(* IEC 61131-3 sources: Versio-VersionControlSystem/fixtures/projects/TC3_PlcSample_reStrText/TC3_PlcSample_reStrText/LibraryDocumentationSample Project/LibPOUs/B_DocuElements/Note elements, 2 files *)

(* ---- FB_Libdoc_GenericNotes.st ---- *)
(*
.. admonition:: And, by the way...

   You can make up your own admonition too.
*)

FUNCTION_BLOCK FB_Libdoc_GenericNotes
VAR_INPUT
    nVarA : INT;
    nVarB : INT;
END_VAR
VAR_OUTPUT
    nSum : INT;
END_VAR
VAR
END_VAR

(* ---- FB_Libdoc_SpecificNotes.st ---- *)
(*
.. note:: This is a note admonition.
   This is the second line of the first paragraph.

   - The note contains all indented body elements
     following.
   - It includes this bullet list.
*)

FUNCTION_BLOCK FB_Libdoc_SpecificNotes
VAR_INPUT
    nVarA : INT;
    nVarB : INT;
END_VAR
VAR_OUTPUT
    nSum : INT;
END_VAR
VAR
END_VAR
